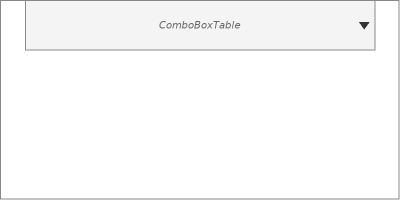
VISUALIZATION V_GCode  // 400x200
VAR_IN_OUT
    HMI_Loader : ST_UsbGcodeLoader_HMI;
END_VAR
    ComboBoxTable (25,0 350x50), variable: HMI_Loader.iSelectedFile, data array: HMI_Loader.aFileList
        p3854506369: HMI_Loader.aFileList[INDEX]
END_VISUALIZATION

(* stored: Version 1.1.0.1, ProductVersion 3.1.4024.15
   Visu V_GCode: Id {db1837f6-f0df-4dac-977b-238054cc0486} *)
